(* PLC project , Example Fixture *)

PROGRAM Calc
  VAR_INPUT
    A : DINT;
  END_VAR
  VAR_OUTPUT
    R : DINT;
  END_VAR
  VAR
    Spent : DINT;
  END_VAR

(* FBD diagram, written out as Structured Text *)
R := A + 1;
END_PROGRAM

CONFIGURATION c
  RESOURCE r ON PLC
  END_RESOURCE
END_CONFIGURATION
